TYPE U_MOVER_SELECTOR_CTRL :
UNION
  stCtrl              : ST_MOVER_SELECTOR_CTRL;

  byCtrl    AT %Q*    : ARRAY[1..SIZEOF(ST_MOVER_SELECTOR_CTRL)] OF BYTE;

END_UNION
END_TYPE

(* stored: Version 1.1.0.1
   DUT U_MOVER_SELECTOR_CTRL: Id {3dae2c87-ee88-480d-ac3a-fb453a81373c} *)
